// TIA Portal V21 export
TagTable "T_V7"
  Y_V7 :   (PLC tag HMI_IF.SwOn, HMI_Connection_1, 1 s)
